SUBAPPLICATION AX_SoftkeyAuxToggle_TO_QXA_BG (* SoftKey (Loslassen) ODER AUX kippt ein Toggle-Flip-Flop (AX_T_FF) auf QXA, Hintergrund SoftKey+AUX spiegelt den Zustand *)
  (* Standard: 61499-2; Description: Copyright (c) 2026 Meisterschulen am Ostbahnhof This program and the accompanying materials are made available under the terms of the Eclipse Public License 2.0 which is available at https://www.eclipse.org/legal/epl-2.0/ SPDX-License-Identifier: EPL-2.0 *)
  (* Version 1.0, 2026-10-31, Franz Höpfinger, Meisterschulen am Ostbahnhof, Aus Getreidehacke func/Manual/Working_Light in MyLib::sys verschoben und umbenannt, INIT/INITO/QI/QO ergaenzt, Output als Parameter (vorher fest Output_Q1). Wie AX_SoftkeyToggle_TO_QXA_BG, zusaetzlich AUX. *)
  PACKAGE MyLib::sys;
  IMPORT isobus::UT::Q::const::IDs::ID_NULL;
  IMPORT logiBUS::io::DQ::logiBUS_DO;
  IMPORT logiBUS::io::DQ::logiBUS_DO_S;
  IMPORT isobus::UT::io::Softkey::SoftKeyActivationCode::SK_RELEASED;
  IMPORT isobus::UT::io::Auxiliary::IN::AuxiliaryState::AuxDisabled_START;
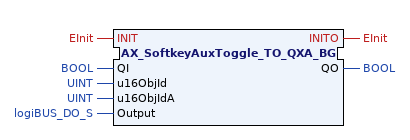
  EVENT_INPUT
    INIT : EInit; (* Initialization Request *)
  END_EVENT
  EVENT_OUTPUT
    INITO : EInit; (* Initialization Confirm *)
  END_EVENT
  VAR_INPUT
    QI : BOOL := TRUE; (* Quality Input - TRUE to enable service *)
    u16ObjId : UINT := ID_NULL; (* Object ID SoftKey *)
    u16ObjIdA : UINT := ID_NULL; (* Object ID AuxFunction2 *)
    Output : logiBUS::io::DQ::logiBUS_DO_S := logiBUS_DO::Invalid; (* logiBUS-Ausgang *)
  END_VAR
  VAR_OUTPUT
    QO : BOOL; (* Quality Output - TRUE if service executed successfully *)
  END_VAR
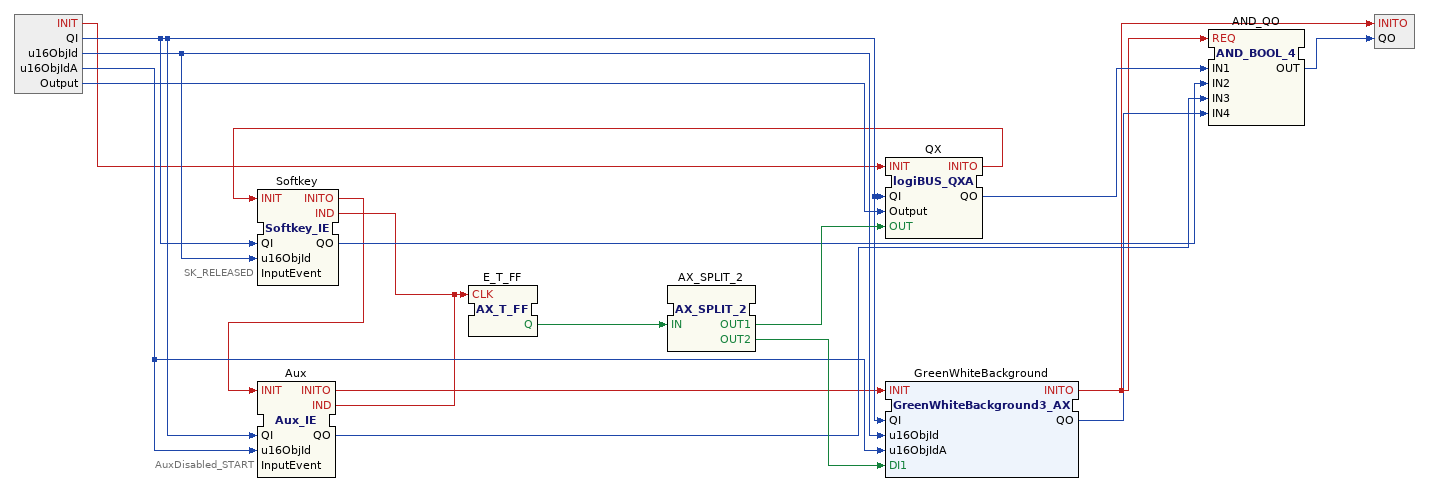
  FBS
    Softkey : isobus::UT::io::Softkey::Softkey_IE(InputEvent := SK_RELEASED);
    Aux : isobus::UT::io::Auxiliary::IN::Aux_IE(InputEvent := AuxDisabled_START);
    E_T_FF : adapter::events::unidirectional::AX_T_FF;
    AX_SPLIT_2 : adapter::events::unidirectional::AX_SPLIT_2;
    QX : logiBUS::io::DQ::logiBUS_QXA;
    AND_QO : iec61131::booleanOperators::AND_BOOL_4;
  END_FBS
  SUBAPPS
    GreenWhiteBackground : MyLib::sys::GreenWhiteBackground3_AX;
  END_SUBAPPS
  EVENT_CONNECTIONS
    INIT TO QX.INIT;
    QX.INITO TO Softkey.INIT;
    Softkey.INITO TO Aux.INIT;
    Aux.INITO TO GreenWhiteBackground.INIT;
    GreenWhiteBackground.INITO TO INITO;
    GreenWhiteBackground.INITO TO AND_QO.REQ;
    Softkey.IND TO E_T_FF.CLK;
    Aux.IND TO E_T_FF.CLK;
  END_CONNECTIONS
  DATA_CONNECTIONS
    QI TO QX.QI;
    QI TO Softkey.QI;
    QI TO Aux.QI;
    QI TO GreenWhiteBackground.QI;
    u16ObjId TO Softkey.u16ObjId;
    u16ObjIdA TO Aux.u16ObjId;
    u16ObjId TO GreenWhiteBackground.u16ObjId;
    u16ObjIdA TO GreenWhiteBackground.u16ObjIdA;
    Output TO QX.Output;
    QX.QO TO AND_QO.IN1;
    Softkey.QO TO AND_QO.IN2;
    Aux.QO TO AND_QO.IN3;
    GreenWhiteBackground.QO TO AND_QO.IN4;
    AND_QO.OUT TO QO;
  END_CONNECTIONS
  ADAPTER_CONNECTIONS
    E_T_FF.Q TO AX_SPLIT_2.IN;
    AX_SPLIT_2.OUT1 TO QX.OUT;
    AX_SPLIT_2.OUT2 TO GreenWhiteBackground.DI1;
  END_CONNECTIONS
END_SUBAPPLICATION
